{attribute 'qualified_only'}
{attribute 'strict'}
TYPE E_CmControlModuleState :
(
	NoCmd
);
END_TYPE

(* stored: Version 1.1.0.1, ProductVersion 3.1.4024.12
   DUT E_CmControlModuleState: Id {f6a7afa2-6b46-4811-b391-ff4c789537f5} *)
